(* IEC 61131-3 sources: RootPLC/conformance/cases/stdlib, 33 files *)

(* ---- err_sizeof_fb.st ---- *)
(* spec: [stdlib.compat.sizeof]
   libraries: TwinCAT_BuiltIns
   expect: error RP0121 *)
FUNCTION_BLOCK FB_X
VAR
    n : INT;
END_VAR
END_FUNCTION_BLOCK

PROGRAM PRG_Main
VAR
    fb : FB_X;
    n : UDINT;
END_VAR
n := SIZEOF(fb);
END_PROGRAM

(* ---- ok_compat_dynamic.st ---- *)
(* spec: [stdlib.compat.dynamic]
   libraries: TwinCAT_BuiltIns
   expect: warning RP0006
   run: PRG_Main cycles=1
   assert: a = 42
   assert: b = 7
   assert: gone = TRUE *)
FUNCTION_BLOCK FB_Node
VAR_INPUT
    v : INT;
END_VAR
METHOD Get : INT
Get := v;
END_METHOD
END_FUNCTION_BLOCK

PROGRAM PRG_Main
VAR
    p : REF_TO INT;
    f : REF_TO FB_Node;
    a, b : INT;
    gone : BOOL;
END_VAR
p := __NEW(INT);
p^ := 41;
a := p^ + 1;
f := __NEW(FB_Node);
f^.v := 7;
b := f^.Get();
__DELETE(p);
__DELETE(f);
gone := p = NULL AND f = NULL;
END_PROGRAM

(* ---- ok_compat_intrinsics.st ---- *)
(* spec: [stdlib.compat.intrinsics]
   libraries: TwinCAT_BuiltIns
   expect: warning RP0006
   run: PRG_Main cycles=3
   assert: who = 'FB_Who'
   assert: t >= T#0MS *)
FUNCTION_BLOCK FB_Who
VAR_OUTPUT
    name : STRING;
END_VAR
name := __POUNAME();
END_FUNCTION_BLOCK

PROGRAM PRG_Main
VAR
    f : FB_Who;
    who : STRING;
    t : TIME;
END_VAR
f();
who := f.name;
t := TIME();
END_PROGRAM

(* ---- ok_compat_query.st ---- *)
(* spec: [stdlib.compat.query]
   libraries: TwinCAT_BuiltIns
   expect: warning RP0006
   run: PRG_Main cycles=1
   assert: hasExtra = TRUE
   assert: noExtra = FALSE
   assert: v = 42
   assert: gotPointer = TRUE *)
INTERFACE I_Base
METHOD Name : INT
END_METHOD
END_INTERFACE

INTERFACE I_Extra
METHOD Extra : INT
END_METHOD
END_INTERFACE

FUNCTION_BLOCK FB_A IMPLEMENTS I_Base, I_Extra
METHOD Name : INT
Name := 1;
END_METHOD
METHOD Extra : INT
Extra := 42;
END_METHOD
END_FUNCTION_BLOCK

FUNCTION_BLOCK FB_B IMPLEMENTS I_Base
METHOD Name : INT
Name := 2;
END_METHOD
END_FUNCTION_BLOCK

PROGRAM PRG_Main
VAR
    a : FB_A;
    b : FB_B;
    ib : I_Base;
    ie : I_Extra;
    p : REF_TO FB_A;
    hasExtra, noExtra, gotPointer : BOOL;
    v : INT;
END_VAR
ib := a;
hasExtra := __QUERYINTERFACE(ib, ie);
IF hasExtra THEN
    v := ie.Extra();
END_IF;
ib := b;
noExtra := __QUERYINTERFACE(ib, ie);
gotPointer := __QUERYPOINTER(a, p);
END_PROGRAM

(* ---- ok_sizeof_array_bound.st ---- *)
(* spec: [variables.constant-names] [stdlib.compat.sizeof]
   libraries: TwinCAT_BuiltIns
   expect: ok
   run: PRG_Main cycles=1
   assert: a = 16
   assert: b = 15
   assert: c = 8
   assert: d = 16 *)
TYPE ST_Cmd :
STRUCT
    id : UINT;
    value : LREAL;
END_STRUCT;
END_TYPE

FUNCTION_BLOCK FB_Sender
VAR
    _command : ST_Cmd;
END_VAR
METHOD PayloadSize : DINT
VAR
    payload : ARRAY[1..SIZEOF(_command)] OF BYTE;
END_VAR
PayloadSize := UPPER_BOUND(payload, 1);
END_METHOD
END_FUNCTION_BLOCK

PROGRAM PRG_Main
VAR
    cmd : ST_Cmd;
    raw : ARRAY[1..SIZEOF(cmd)] OF BYTE;
    raw2 : ARRAY[0..SIZEOF(ST_Cmd) - 1] OF BYTE;
    words : ARRAY[1..SIZEOF(cmd) / SIZEOF(WORD)] OF WORD;
    sender : FB_Sender;
    a, b, c, d : DINT;
END_VAR
a := UPPER_BOUND(raw, 1);
b := UPPER_BOUND(raw2, 1);
c := UPPER_BOUND(words, 1);
d := sender.PayloadSize();
END_PROGRAM

(* ---- ok_tcunit_suite.st ---- *)
(* spec: [stdlib.compat.unit]
   libraries: TcUnit
   expect: ok
   run: PRG_TEST cycles=10 *)
FUNCTION_BLOCK FB_CounterTests EXTENDS FB_TestSuite
Increments();
Wraps();
METHOD Increments
VAR
    n : INT := 41;
END_VAR
TEST('Increments');
n := n + 1;
AssertEquals_INT(Expected := 42, Actual := n, Message := 'one more');
TEST_FINISHED();
END_METHOD
METHOD Wraps
VAR
    b : USINT := 255;
END_VAR
TEST('Wraps');
b := b + 1;
AssertEquals(Expected := USINT#0, Actual := b, Message := 'USINT wraps');
AssertTrue(Condition := b = 0, Message := 'zero');
TEST_FINISHED();
END_METHOD
END_FUNCTION_BLOCK

PROGRAM PRG_TEST
VAR
    counter : FB_CounterTests;
END_VAR
TcUnit.RUN();
END_PROGRAM

(* ---- warn_compat_eventlogger.st ---- *)
(* spec: [stdlib.compat.declare-only]
   libraries: Tc3_EventLogger
   expect: warning RP0118 RP0120
   run: PRG_Main cycles=1
   assert: n = 7
   assert: ok = TRUE
   assert: same = TRUE
   assert: sev = TcEventSeverity#Warning *)
FUNCTION_BLOCK FB_Listener EXTENDS FB_ListenerBase2
VAR
    nMessages : UDINT;
END_VAR
METHOD OnMessageSent : HRESULT
VAR_INPUT
    fbEvent : REFERENCE TO FB_TcEvent;
END_VAR
nMessages := nMessages + 1;
END_METHOD
END_FUNCTION_BLOCK

PROGRAM PRG_Main
VAR
    send : BOOL;
    fbMsg : FB_TcMessage;
    fbAlarm : FB_TcAlarm;
    listener : FB_Listener;
    entry : TcEventEntry;
    src, other : FB_TcSourceInfo;
    ipSrc : I_TcSourceInfo := NULL;
    hr : HRESULT;
    ok, same : BOOL;
    n : UDINT;
    sev : TcEventSeverity;
END_VAR
src.sName := 'Main';
ok := src.ExtendName('.Pump');
src.nId := 7;
other.sName := 'Main.Pump';
other.nId := 7;
ipSrc := other;
same := src.EqualsTo(ipSrc);
n := src.nId;
entry.eSeverity := TcEventSeverity#Warning;
sev := entry.eSeverity;
IF send THEN
    (* declared only: a run that reaches these stops with UNSUPPORTED *)
    hr := fbMsg.CreateEx(entry, src);
    fbMsg.ipArguments.Clear().AddString('pump').AddInt(3);
    hr := fbMsg.Send(0);
    IF fbAlarm.bRaised THEN
        hr := fbAlarm.Clear(0, FALSE);
    END_IF;
    hr := listener.Execute();
END_IF;
END_PROGRAM

(* ---- compat_ads_error_enums.st ---- *)
(* spec: [stdlib.compat]
   libraries: Tc2_System
   expect: warning RP0122 RP0129
   run: PRG_Main cycles=1
   assert: n = 2
   assert: code = 1802
   assert: hr = -1743714549
   assert: failed = TRUE *)
FUNCTION F_Check : HRESULT
VAR_INPUT
    n : INT;
END_VAR
IF n < 0 THEN
    F_Check := Tc2_System.E_HRESULTAdsErr.INVALIDPARM;
ELSE
    F_Check := E_HRESULTAdsErr.HRESULT_ADS_NOERROR;
END_IF;
END_FUNCTION

PROGRAM PRG_Main
VAR
    hr : HRESULT;
    e : E_AdsErr;
    n : INT;
    code : UDINT;
    failed : BOOL;
END_VAR
hr := F_Check(-1);
CASE hr OF
    E_HRESULTAdsErr.HRESULT_ADS_NOERROR: n := 1;
    E_HRESULTAdsErr.INVALIDPARM: n := 2;
END_CASE;
e := E_AdsErr.DEVICE_NOMEMORY;
IF e <> E_AdsErr.NOERR THEN
    code := e;
END_IF;
failed := hr < 0;
END_PROGRAM

(* ---- compat_json_sax_writer.st ---- *)
(* spec: [stdlib.compat]
   libraries: Tc3_JsonXml
   expect: ok
   run: PRG_Main cycles=1
   assert: sDoc = '{"Timestamp":"2017-04-04T12:42:42","Values":{"Sensor2":[1,2,-3],"On":true,"Name":"Pump \"A\"\\1","Off":null},"Raw":{"x":42},"Big":18446744073709551615}'
   assert: nLen = 151
   assert: nCopied = 152
   assert: sCopy = '{"Timestamp":"2017-04-04T12:42:42","Values":{"Sensor2":[1,2,-3],"On":true,"Name":"Pump \"A\"\\1","Off":null},"Raw":{"x":42},"Big":18446744073709551615}'
   assert: nTooSmall = 0
   assert: sSmall = ''
   assert: sAfterReset = '[]' *)
PROGRAM PRG_Main
VAR
    fbJson : FB_JsonSaxWriter;
    dtTimestamp : DT := DT#2017-04-04-12:42:42;
    sDoc : STRING[255];
    sCopy : STRING[1000];
    sSmall : STRING[10] := 'old';
    sAfterReset : STRING[255];
    nLen, nCopied, nTooSmall : UDINT;
END_VAR
fbJson.ResetDocument();
fbJson.StartObject();
fbJson.AddKeyDateTime('Timestamp', dtTimestamp);
fbJson.AddKey('Values');
fbJson.StartObject();
fbJson.AddKey('Sensor2');
fbJson.StartArray();
fbJson.AddDint(1);
fbJson.AddUdint(2);
fbJson.AddLint(-3);
fbJson.EndArray();
fbJson.AddKeyBool('On', TRUE);
fbJson.AddKeyString('Name', 'Pump "A"\1');
fbJson.AddKeyNull('Off');
fbJson.EndObject();
fbJson.AddKey('Raw');
fbJson.AddRawObject('{"x":42}');
fbJson.AddKey('Big');
fbJson.AddUlint(18446744073709551615);
fbJson.EndObject();
sDoc := fbJson.GetDocument();
nLen := fbJson.GetDocumentLength();
nCopied := fbJson.CopyDocument(sCopy, SIZEOF(sCopy));
nTooSmall := fbJson.CopyDocument(sSmall, SIZEOF(sSmall));
fbJson.ResetDocument();
fbJson.StartArray();
fbJson.EndArray();
sAfterReset := fbJson.GetDocument();
END_PROGRAM

(* ---- err_fb_input_type.st ---- *)
(* spec: [stdlib.fbs]
   expect: error RP0103 *)
PROGRAM PRG_Main
VAR
    t : TON;
END_VAR
t(IN := TRUE, PT := 500);
END_PROGRAM

(* ---- err_no_common_type.st ---- *)
(* spec: [stdlib.functions]
   expect: error RP0103 *)
PROGRAM PRG_Main
VAR
    i : INT;
    b : BOOL;
END_VAR
i := MAX(i, b);
END_PROGRAM

(* ---- ok_compat_adslog.st ---- *)
(* spec: [stdlib.compat.log]
   libraries: Tc2_System
   expect: ok
   run: PRG_Main cycles=2
   assert: res = 0
   assert: count = 2 *)
PROGRAM PRG_Main
VAR
    res : DINT := -1;
    count : DINT;
END_VAR
count := count + 1;
res := ADSLOGSTR(ADSLOG_MSGTYPE_HINT, 'Started %s', 'motor');
res := res + ADSLOGDINT(ADSLOG_MSGTYPE_WARN, 'Cycle %d', count);
res := res + ADSLOGLREAL(ADSLOG_MSGTYPE_ERROR, 'Speed %f', 1.5);
END_PROGRAM

(* ---- ok_compat_any.st ---- *)
(* spec: [stdlib.compat.any]
   libraries: TwinCAT_BuiltIns
   expect: warning RP0006 RP0122
   run: PRG_Main cycles=1
   assert: a = 702
   assert: b = -15
   assert: c = 502 *)
FUNCTION F_Describe : DINT
VAR_INPUT
    value : ANY;
END_VAR
VAR
    pI : REF_TO INT;
END_VAR
IF value.TypeClass = __SYSTEM.TYPE_CLASS.TYPE_INT THEN
    pI := value.pValue;
    F_Describe := INT_TO_DINT(pI^) * 100 + value.diSize;
ELSE
    F_Describe := -TO_DINT(value.TypeClass);
END_IF;
END_FUNCTION

PROGRAM PRG_Main
VAR
    i : INT := 7;
    r : LREAL := 1.0;
    a, b, c : DINT;
END_VAR
a := F_Describe(i);
b := F_Describe(r);
c := F_Describe(INT#5);
END_PROGRAM

(* ---- ok_compat_clock.st ---- *)
(* spec: [stdlib.compat.clock]
   libraries: Tc2_System
   expect: ok
   run: PRG_Main cycles=2
   assert: first = ULINT#134116992000000000
   assert: now = first *)
(* The virtual time of day starts at 2026-01-01 00:00:00 UTC (a file time
   in 100 ns units); the conformance runner does not advance the clock. *)
PROGRAM PRG_Main
VAR
    first : ULINT;
    now : ULINT;
END_VAR
IF first = 0 THEN
    first := F_GetSystemTime();
END_IF;
now := F_GetSystemTime();
END_PROGRAM

(* ---- ok_compat_formatstring.st ---- *)
(* spec: [stdlib.compat]
   libraries: Tc2_Utilities
   expect: ok
   run: PRG_Main cycles=1
   assert: measure = 'Measure X: +0000000130, Y: +0000000130'
   assert: ints = '-5|   -5|-5   |'
   assert: bits = 'ab AB 16#ab 10101011 454'
   assert: reals = '3.141590|3.14|+003.142|-2.500000'
   assert: strs = '[hello] [hel] [   hello] [hello   ] 100%'
   assert: misc = 'A42       -5 ff'
   assert: missing = 16386
   assert: badType = 2049
   assert: mismatch = 4097
   assert: failed = TRUE *)
PROGRAM PRG_Main
VAR
    fmt, fresh1, fresh2, fresh3 : FB_FormatString;
    x : DINT := 130;
    neg : INT := -5;
    b : BYTE := 16#AB;
    w : WORD := 300;
    r : LREAL := 3.14159;
    rr : REAL := -2.5;
    s : T_MaxString := 'hello';
    u : UDINT := 42;
    ch : BYTE := 65;
    wd : UDINT := 8;
    sb : SINT := -1;
    measure, ints, bits, reals, strs, misc : T_MaxString;
    missing, badType, mismatch : UDINT;
    failed : BOOL;
END_VAR
fmt(sFormat := 'Measure X: %+.10d, Y: %+.10d', arg1 := F_DINT(x), arg2 := F_DINT(x));
measure := fmt.sOut;
fmt(sFormat := '%d|%5d|%-5d|', arg1 := F_INT(neg), arg2 := F_INT(neg), arg3 := F_INT(neg));
ints := fmt.sOut;
fmt(sFormat := '%x %X %#x %b %o', arg1 := F_BYTE(b), arg2 := F_BYTE(b), arg3 := F_BYTE(b),
    arg4 := F_BYTE(b), arg5 := F_WORD(w));
bits := fmt.sOut;
fmt(sFormat := '%f|%.2f|%+08.3f|%f', arg1 := F_LREAL(r), arg2 := F_LREAL(r), arg3 := F_LREAL(r),
    arg4 := F_REAL(rr));
reals := fmt.sOut;
fmt(sFormat := '[%s] [%.3s] [%8s] [%-8s] 100%%', arg1 := F_STRING(s), arg2 := F_STRING(s),
    arg3 := F_STRING(s), arg4 := F_STRING(s));
strs := fmt.sOut;
fmt(sFormat := '%c%u %*d %x', arg1 := F_BYTE(ch), arg2 := F_UDINT(u), arg3 := F_INT(neg),
    arg4 := F_UDINT(wd), arg5 := F_SINT(sb));
misc := fmt.sOut;
fresh1(sFormat := '%d %d', arg1 := F_INT(neg));
missing := fresh1.nErrId;
failed := fresh1.bError;
fresh2(sFormat := '%q', arg1 := F_INT(neg));
badType := fresh2.nErrId;
fresh3(sFormat := '%s', arg1 := F_INT(neg));
mismatch := fresh3.nErrId;
END_PROGRAM

(* ---- ok_compat_hexstr.st ---- *)
(* spec: [stdlib.compat]
   libraries: Tc2_Utilities
   expect: ok
   run: PRG_Main cycles=1
   assert: a = 'FF'
   assert: b = '000f'
   assert: c = ''
   assert: d = 'ABCD'
   assert: e = '0' *)
PROGRAM PRG_Main
VAR
    a, b, c, d, e : T_MaxString;
END_VAR
a := BYTE_TO_HEXSTR(16#FF, 1, FALSE);
b := WORD_TO_HEXSTR(15, 4, TRUE);
c := DWORD_TO_HEXSTR(0, 0, FALSE);
d := LWORD_TO_HEXSTR(43981, 1, FALSE);
e := BYTE_TO_HEXSTR(0, 1, FALSE);
END_PROGRAM

(* ---- ok_compat_tc2_standard.st ---- *)
(* spec: [stdlib.compat]
   libraries: Tc2_Standard
   expect: ok
   run: PRG_Main cycles=3
   assert: n = 4
   assert: m = "US"
   assert: s = "SUSIX"
   assert: f = 0
   assert: up = 2
   assert: hit = TRUE
   assert: down = 4
   assert: both = 0
   assert: pulse = TRUE
   assert: off = TRUE *)
PROGRAM PRG_Main
VAR
    n, f : INT;
    m, s : WSTRING;
    clk : BOOL;
    hit, pulse, off : BOOL;
    up, down, both : WORD;
    cu : CTU;
    cd : CTD;
    cud : CTUD;
    lp : LTP;
    lf : LTOF;
END_VAR
n := WLEN("SUSI");
m := WMID("SUSI", 2, 2);
s := WCONCAT("SUSI", "X");
f := WFIND("SUSI", "Q");
clk := NOT clk;
cu(CU := clk, RESET := FALSE, PV := 2);
up := cu.CV;
hit := cu.Q;
cd(CD := FALSE, LOAD := TRUE, PV := 4);
down := cd.CV;
cud(CU := clk, CD := FALSE, RESET := TRUE, LOAD := FALSE, PV := 5);
both := cud.CV;
lp(IN := TRUE, PT := LTIME#1S);
pulse := lp.Q;
lf(IN := TRUE, PT := LTIME#1S);
off := lf.Q;
END_PROGRAM

(* ---- ok_compat_tc2_system.st ---- *)
(* spec: [stdlib.compat]
   libraries: Tc2_System, TwinCAT_BuiltIns
   expect: ok
   run: PRG_Main cycles=1
   assert: n = 255
   assert: r > 6.28 AND r < 6.29
   assert: ready *)
TYPE ST_Flags : STRUCT
    running : BIT;
END_STRUCT; END_TYPE

PROGRAM PRG_Main
VAR
    s : T_MaxString := 'motor';
    n : UDINT;
    r : LREAL;
    f : ST_Flags;
    ready : BOOL;
END_VAR
n := MAX_STRING_LENGTH;
r := Tc2_System.PI * 2.0;
f.running := ADSLOG_MSGTYPE_HINT = 16#01;
ready := f.running;
END_PROGRAM

(* ---- ok_compat_tc2_system_info.st ---- *)
(* spec: [stdlib.compat]
   libraries: Tc2_System, TwinCAT_BuiltIns
   expect: warning RP0006 RP0122
   run: PRG_Main cycles=1
   assert: older = -1
   assert: same = 0
   assert: taskNo = 1
   assert: idx = 1
   assert: cls = TRUE
   assert: port = 851 *)
PROGRAM PRG_Main
VAR
    v : ST_LibVersion := (iMajor := 3, iMinor := 4, iBuild := 1, iRevision := 0);
    older, same, idx : DINT;
    taskNo : BYTE;
    getIdx : GETCURTASKINDEX;
    tc : __SYSTEM.TYPE_CLASS;
    cls : BOOL;
    addr : ST_AmsAddr;
    port : UINT;
    first : BOOL;
END_VAR
older := F_CmpLibVersion(v, 3, 5, 0, 0);
same := F_CmpLibVersion(v, 3, 4, 1, 0);
getIdx();
taskNo := getIdx.index;
idx := GETCURTASKINDEXEX();
first := TwinCAT_SystemInfoVarList._TaskInfo[idx].FirstCycle;
tc := __SYSTEM.TYPE_CLASS.TYPE_LREAL;
cls := TO_DWORD(tc) = 15;
addr.port := 851;
port := addr.port;
END_PROGRAM

(* ---- ok_compat_tc2_utilities_strings.st ---- *)
(* spec: [stdlib.compat]
   libraries: Tc2_Utilities
   expect: ok
   run: PRG_Main cycles=1
   assert: lower = 'to lower case 1234567890 äöüß'
   assert: upper = 'ABC ÄÖ'
   assert: left = '<trim '
   assert: right = ' trim>'
   assert: kind = TRUE
   assert: size = 4 *)
PROGRAM PRG_Main
VAR
    lower, upper, left, right : T_MaxString;
    value : DINT := 7;
    arg : T_Arg;
    kind : BOOL;
    size : UDINT;
    stamp : TIMESTRUCT;
END_VAR
lower := F_ToLCase('TO LOWER CASE 1234567890 ÄÖÜß');
upper := F_ToUCase('abc äö');
left := F_LTrim(' <trim ');
right := F_RTrim(' trim> ');
arg := F_DINT(value);
kind := arg.eType = E_ArgType#ARGTYPE_DINT;
size := arg.cbLen;
stamp.wYear := 2026;
END_PROGRAM

(* ---- ok_compat_tc2_utilities_time.st ---- *)
(* spec: [stdlib.compat]
   libraries: Tc2_Utilities
   expect: warning RP0117
   run: PRG_Main cycles=1
   assert: text = '2026-11-04-12:30:15.000'
   assert: weekday = 3
   assert: back = TRUE
   assert: ft = 134382690150000000
   assert: rounded = '0.47'
   assert: cut = '0.46'
   assert: copied = 'hel'
   assert: complete = FALSE
   assert: netId = '127.16.17.3.1.1' *)
PROGRAM PRG_Main
VAR
    stamp : DT := DT#2026-11-04-12:30:15;
    st : TIMESTRUCT;
    text : STRING;
    weekday : WORD;
    back : BOOL;
    ft : T_FILETIME64;
    rounded, cut : STRING[510];
    src : STRING := 'hello';
    copied : STRING;
    complete : BOOL;
    ids : T_AmsNetIdArr := [127, 16, 17, 3, 1, 1];
    netId : T_AmsNetId;
END_VAR
st := DT_TO_SYSTEMTIME(stamp);
text := SYSTEMTIME_TO_STRING(st);
weekday := st.wDayOfWeek;
back := SYSTEMTIME_TO_DT(st) = stamp;
ft := SYSTEMTIME_TO_FILETIME64(st);
rounded := LREAL_TO_FMTSTR(0.46523, 2, TRUE);
cut := LREAL_TO_FMTSTR(0.46523, 2, FALSE);
complete := STRNCPY(ADR(copied), ADR(src), 4);
netId := F_CreateAmsNetId(ids);
END_PROGRAM

(* ---- ok_compat_tc3_module.st ---- *)
(* spec: [stdlib.compat]
   libraries: Tc3_Module
   expect: ok
   run: PRG_Main cycles=1
   assert: ok = TRUE
   assert: bad = TRUE
   assert: pending = 515 *)
PROGRAM PRG_Main
VAR
    hr : HRESULT := S_OK;
    ok, bad : BOOL;
    pending : DINT;
END_VAR
ok := SUCCEEDED(hr) AND SUCCEEDED(S_FALSE);
hr := -2147467259;
bad := FAILED(hr);
pending := S_PENDING;
END_PROGRAM

(* ---- ok_functions.st ---- *)
(* spec: [stdlib.conversions] [stdlib.functions]
   expect: ok
   run: PRG_Main cycles=1
   assert: d = 2
   assert: i = 3
   assert: w = 16#0F00
   assert: n = 4 *)
PROGRAM PRG_Main
VAR
    i : INT := -7;
    d : DINT;
    r : LREAL := 2.7;
    w : WORD := 16#00F0;
    s : STRING;
    n : INT;
END_VAR
d := INT_TO_DINT(ABS(i));
d := TRUNC(r);
i := LIMIT(0, i, 100);
i := MAX(i, 3);
w := SHL(w, 4);
s := CONCAT('ab', 'cd');
n := LEN(s);
r := TO_LREAL(n) + SQRT(r);
END_PROGRAM

(* ---- ok_open_array_bounds.st ---- *)
(* spec: [stdlib.functions.bounds]
   expect: ok
   run: PRG_Main cycles=1
   assert: s1 = 6
   assert: s2 = 30
   assert: lo = 2
   assert: hi = 4
   assert: x[3] = 0
   assert: m = 20 *)
FUNCTION SumAndClear : DINT
VAR_IN_OUT
    a : ARRAY[*] OF INT;
END_VAR
VAR
    i : DINT;
END_VAR
FOR i := LOWER_BOUND(a, 1) TO UPPER_BOUND(a, 1) DO
    SumAndClear := SumAndClear + a[i];
    a[i] := 0;
END_FOR;
END_FUNCTION

FUNCTION MaxOf : INT
VAR_INPUT
    a : ARRAY[*] OF INT;
END_VAR
VAR
    i : DINT;
END_VAR
MaxOf := a[LOWER_BOUND(a, 1)];
FOR i := LOWER_BOUND(a, 1) + 1 TO UPPER_BOUND(a, 1) DO
    MaxOf := MAX(MaxOf, a[i]);
END_FOR;
END_FUNCTION

PROGRAM PRG_Main
VAR
    x : ARRAY[2..4] OF INT := [1, 2, 3];
    y : ARRAY[0..1] OF INT := [10, 20];
    s1, s2, lo, hi : DINT;
    m : INT;
END_VAR
m := MaxOf(y);
s1 := SumAndClear(x);
s2 := SumAndClear(y);
lo := LOWER_BOUND(x, 1);
hi := UPPER_BOUND(x, 1);
END_PROGRAM

(* ---- ok_operator_functions.st ---- *)
(* spec: [stdlib.functions.operators]
   expect: ok
   run: PRG_Main cycles=1
   assert: a = 10
   assert: s = 3
   assert: m = 24
   assert: q = 2
   assert: r = 1
   assert: up = TRUE
   assert: neq = FALSE
   assert: t = T#1500ms *)
PROGRAM PRG_Main
VAR
    a, s, m, q, r : INT;
    up, neq : BOOL;
    t : TIME;
END_VAR
a := ADD(1, 2, 3, 4);
s := SUB(IN1 := 5, IN2 := 2);
m := MUL(2, 3, 4);
q := DIV(7, 3);
r := MOD(7, 3);
up := GT(5, 3, 1) AND LE(1, 1, 2);
neq := NE(4, 4);
t := ADD(T#1S, T#500MS);
END_PROGRAM

(* ---- ok_sizeof.st ---- *)
(* spec: [stdlib.compat.sizeof]
   libraries: TwinCAT_BuiltIns
   expect: warning RP0115
   run: PRG_Main cycles=1
   assert: a = 2
   assert: b = 16
   assert: c = 11
   assert: d = 8
   assert: e = 24
   assert: f = 4
   assert: g = 16 *)
TYPE
    ST_Pair : STRUCT
        dw : DWORD;
        lw : LWORD;
    END_STRUCT;
    ST_Mixed : STRUCT
        flag : BOOL;
        value : LREAL;
        n : INT;
    END_STRUCT;
    E_Mode : UINT (Off, Auto);
    E_Big : (One, Two) DINT;
END_TYPE

PROGRAM PRG_Main
VAR
    p : ST_Pair;
    s : STRING[10];
    arr : ARRAY[1..4] OF INT;
    a : USINT;
    b, c, d, e, f : USINT;
    g : ULINT;
END_VAR
a := SIZEOF(INT);
b := SIZEOF(p);
c := SIZEOF(s);
d := SIZEOF(arr);
e := SIZEOF(ST_Mixed);
f := SIZEOF(E_Big);
g := XSIZEOF(ST_Pair);
END_PROGRAM

(* ---- ok_standard_fbs.st ---- *)
(* spec: [stdlib.fbs]
   expect: ok *)
PROGRAM PRG_Main
VAR
    start, stop : BOOL;
    t : TON;
    edge : R_TRIG;
    cnt : CTU;
    latch : SR;
    count : INT;
    elapsed : TIME;
END_VAR
t(IN := start, PT := T#2s, ET => elapsed);
edge(CLK := start);
cnt(CU := edge.Q, R := stop, PV := 10);
count := cnt.CV;
latch(S1 := t.Q, R := stop);
END_PROGRAM

(* ---- ok_string_result_length.st ---- *)
(* spec: [stdlib.string.length]
   expect: ok
   run: PRG_Main cycles=1
   assert: a = 120
   assert: b = 160
   assert: c = 10
   assert: d = 125 *)
PROGRAM PRG_Main
VAR
    s60 : STRING[60] := '012345678901234567890123456789012345678901234567890123456789';
    long : STRING[300];
    short : STRING[10];
    a, b, c, d : INT;
END_VAR
long := CONCAT(s60, s60);
a := LEN(long);
long := CONCAT(long, CONCAT(s60, LEFT(s60, 40)));
a := LEN(CONCAT(s60, s60));
b := LEN(LEFT(long, 160));
short := CONCAT(s60, 'x');
c := LEN(short);
d := LEN(INSERT(long, 'abcde', 3)) - 100;
END_PROGRAM

(* ---- ok_task_info.st ---- *)
(* spec: [stdlib.compat.taskinfo]
   libraries: TwinCAT_BuiltIns, Tc2_System
   expect: ok *)
PROGRAM PRG_Main
VAR
    cycleMs : UDINT;
END_VAR
cycleMs := _TaskInfo[GETCURTASKINDEXEX()].CycleTime / 10000;
END_PROGRAM

(* ---- warn_compat_declare_only.st ---- *)
(* spec: [stdlib.compat.declare-only]
   libraries: Tc2_System
   expect: warning RP0120
   run: PRG_Main cycles=1
   assert: x = 0.0 *)
PROGRAM PRG_Main
VAR
    draw : BOOL;
    rnd : DRAND;
    x : LREAL;
END_VAR
IF draw THEN
    rnd(Seed := 1);
    x := rnd.Num;
END_IF;
END_PROGRAM

(* ---- warn_compat_json_declare_only.st ---- *)
(* spec: [stdlib.compat.declare-only]
   libraries: Tc3_JsonXml
   expect: warning RP0120
   run: PRG_Main cycles=1
   assert: n = 2 *)
PROGRAM PRG_Main
VAR
    parse : BOOL;
    fbDom : FB_JsonDomParser;
    fbJson : FB_JsonSaxWriter;
    jsonDoc, jsonProp : SJsonValue;
    sDoc : STRING[255] := '{"a":1}';
    f : LREAL;
    n : UDINT;
END_VAR
fbJson.StartArray();
fbJson.AddDint(1);
IF parse THEN
    (* declared only: a run that reaches these stops with UNSUPPORTED *)
    jsonDoc := fbDom.ParseDocument(sDoc);
    jsonProp := fbDom.FindMember(jsonDoc, 'a');
    f := fbDom.GetDouble(jsonProp);
    fbJson.AddLreal(f);
END_IF;
fbJson.EndArray();
n := fbJson.GetDocumentLength() - 1;
END_PROGRAM

(* ---- warn_compat_memcpy.st ---- *)
(* spec: [stdlib.compat.pvoid]
   libraries: Tc2_System
   expect: warning RP0117 RP0120 *)
PROGRAM PRG_Main
VAR
    a, b : ARRAY[0..3] OF INT;
    p : PVOID;
    n : UDINT;
    same : DINT;
END_VAR
p := ADR(a);
n := MEMCPY(destAddr := p, srcAddr := ADR(b), n := SIZEOF(b));
n := MEMSET(ADR(a), 0, SIZEOF(a));
same := MEMCMP(ADR(a), ADR(b), SIZEOF(a));
END_PROGRAM

(* ---- warn_compat_tc2_mc2.st ---- *)
(* spec: [stdlib.compat.declare-only]
   libraries: Tc2_MC2
   expect: warning RP0120 *)
PROGRAM PRG_Main
VAR
    axis : AXIS_REF;
    power : MC_Power;
    move : MC_MoveAbsolute;
    pos : LREAL;
    ready : BOOL;
END_VAR
power(Enable := TRUE, Enable_Positive := TRUE, Enable_Negative := TRUE, Axis := axis);
move(Execute := power.Status, Position := 100.0, Velocity := 50.0, Axis := axis);
axis.ReadStatus();
pos := axis.NcToPlc.ActPos;
ready := axis.Status.StandStill AND NOT axis.Status.Error;
axis.PlcToNc.Override := 100;
END_PROGRAM
